(*
SPDX-FileCopyrightText: © 2026 Oleksandr Tiutyk <trofimich@gmail.com>
SPDX-License-Identifier: MIT
License: https://opensource.org/license/mit
*)

(*!
<summary>Indicates whether a test body needs more scheduling cycles or has finished on the current cycle.</summary>
<description>
BUSY (0) is the default uninitialized value and keeps the test running across subsequent cycles unless a failure
or deadline terminates the run. DONE (1) requests normal completion after the current cycle returns.
</description>
*)

{attribute 'qualified_only'}
{attribute 'strict'}
{attribute 'to_string'}
TYPE TEST_CYCLE_RESULT :
(
	BUSY := 0,
	DONE := 1
);
END_TYPE

(* stored: Version 1.1.0.1
   DUT TEST_CYCLE_RESULT: Id {9cdb4d44-16b2-4bc8-a63b-cd4e52c2f709} *)
